(* IEC 61131-3 sources: crb-codesys/generation/scripts/repoeval/交通信号灯控制实训/global, 3 files *)

(* ---- GVL_Input.st ---- *)
VAR_GLOBAL
	IReset	:	BOOL;
END_VAR

(* ---- GVL_Memory.st ---- *)
VAR_GLOBAL
	MCountBackwards	:	UINT;//剩余时间
	MGreenTimeOn	:	TIME := T#30S;//绿灯亮的时间
	MGreenTimeFlash	:	TIME := T#3S;//绿灯闪的时间
	MYellowTimeOn	:	TIME := T#3S;//黄灯亮的时间
END_VAR

(* ---- GVL_Output.st ---- *)
VAR_GLOBAL
	QSouthNorthGreen	:	BOOL;//与视图中南北方向的绿灯相关联
	QSouthNorthYellow	:	BOOL;
	QSouthNorthRed	:	BOOL;
	QEastWestGreen	:	BOOL;
	QEastWestYellow	:	BOOL;
	QEastWestRed	:	BOOL;
END_VAR
